(* IEC 61131-3 sources: STAR-PLC-Agent/results/raw/four_group_20261114/star_deepseek_v4/SELF011/generation/sim_00, 1 file *)

(* ---- test_program.st ---- *)
PROGRAM PLC_PRG
VAR
 BenchStep : UDINT := 0;
 BenchCalls : UDINT := 0;
 BenchDone : BOOL := FALSE;
 BenchUut0 : FB_Task;
 BenchUut1 : FB_Task;
 TraceIn_Start : ARRAY[0..12] OF BOOL;
 TraceIn_Stop : ARRAY[0..12] OF BOOL;
 TraceIn_Reset : ARRAY[0..12] OF BOOL;
 TraceIn_ExtendDone : ARRAY[0..12] OF BOOL;
 TraceIn_ClampDone : ARRAY[0..12] OF BOOL;
 TraceIn_ReleaseDone : ARRAY[0..12] OF BOOL;
 TraceIn_RetractDone : ARRAY[0..12] OF BOOL;
 TraceOut_Extend : ARRAY[0..12] OF BOOL;
 TraceOut_Clamp : ARRAY[0..12] OF BOOL;
 TraceOut_Release : ARRAY[0..12] OF BOOL;
 TraceOut_Retract : ARRAY[0..12] OF BOOL;
 TraceOut_Busy : ARRAY[0..12] OF BOOL;
 TraceOut_Done : ARRAY[0..12] OF BOOL;
END_VAR

IF NOT BenchDone THEN
 CASE BenchStep OF
 0:
   BenchUut0.Start := TRUE;
   BenchUut0.Stop := FALSE;
   BenchUut0.Reset := FALSE;
   BenchUut0.ExtendDone := FALSE;
   BenchUut0.ClampDone := FALSE;
   BenchUut0.ReleaseDone := FALSE;
   BenchUut0.RetractDone := TRUE;
   TraceIn_Start[0] := BenchUut0.Start;
   TraceIn_Stop[0] := BenchUut0.Stop;
   TraceIn_Reset[0] := BenchUut0.Reset;
   TraceIn_ExtendDone[0] := BenchUut0.ExtendDone;
   TraceIn_ClampDone[0] := BenchUut0.ClampDone;
   TraceIn_ReleaseDone[0] := BenchUut0.ReleaseDone;
   TraceIn_RetractDone[0] := BenchUut0.RetractDone;
   BenchUut0();
   TraceOut_Extend[0] := BenchUut0.Extend;
   TraceOut_Clamp[0] := BenchUut0.Clamp;
   TraceOut_Release[0] := BenchUut0.Release;
   TraceOut_Retract[0] := BenchUut0.Retract;
   TraceOut_Busy[0] := BenchUut0.Busy;
   TraceOut_Done[0] := BenchUut0.Done;
   BenchCalls := BenchCalls + 1;
 1:
   BenchUut0.Start := FALSE;
   BenchUut0.Stop := FALSE;
   BenchUut0.Reset := FALSE;
   BenchUut0.ExtendDone := TRUE;
   BenchUut0.ClampDone := FALSE;
   BenchUut0.ReleaseDone := FALSE;
   BenchUut0.RetractDone := FALSE;
   TraceIn_Start[1] := BenchUut0.Start;
   TraceIn_Stop[1] := BenchUut0.Stop;
   TraceIn_Reset[1] := BenchUut0.Reset;
   TraceIn_ExtendDone[1] := BenchUut0.ExtendDone;
   TraceIn_ClampDone[1] := BenchUut0.ClampDone;
   TraceIn_ReleaseDone[1] := BenchUut0.ReleaseDone;
   TraceIn_RetractDone[1] := BenchUut0.RetractDone;
   BenchUut0();
   TraceOut_Extend[1] := BenchUut0.Extend;
   TraceOut_Clamp[1] := BenchUut0.Clamp;
   TraceOut_Release[1] := BenchUut0.Release;
   TraceOut_Retract[1] := BenchUut0.Retract;
   TraceOut_Busy[1] := BenchUut0.Busy;
   TraceOut_Done[1] := BenchUut0.Done;
   BenchCalls := BenchCalls + 1;
 2:
   BenchUut0.Start := FALSE;
   BenchUut0.Stop := FALSE;
   BenchUut0.Reset := FALSE;
   BenchUut0.ExtendDone := FALSE;
   BenchUut0.ClampDone := TRUE;
   BenchUut0.ReleaseDone := FALSE;
   BenchUut0.RetractDone := FALSE;
   TraceIn_Start[2] := BenchUut0.Start;
   TraceIn_Stop[2] := BenchUut0.Stop;
   TraceIn_Reset[2] := BenchUut0.Reset;
   TraceIn_ExtendDone[2] := BenchUut0.ExtendDone;
   TraceIn_ClampDone[2] := BenchUut0.ClampDone;
   TraceIn_ReleaseDone[2] := BenchUut0.ReleaseDone;
   TraceIn_RetractDone[2] := BenchUut0.RetractDone;
   BenchUut0();
   TraceOut_Extend[2] := BenchUut0.Extend;
   TraceOut_Clamp[2] := BenchUut0.Clamp;
   TraceOut_Release[2] := BenchUut0.Release;
   TraceOut_Retract[2] := BenchUut0.Retract;
   TraceOut_Busy[2] := BenchUut0.Busy;
   TraceOut_Done[2] := BenchUut0.Done;
   BenchCalls := BenchCalls + 1;
 3:
   BenchUut0.Start := FALSE;
   BenchUut0.Stop := FALSE;
   BenchUut0.Reset := FALSE;
   BenchUut0.ExtendDone := FALSE;
   BenchUut0.ClampDone := FALSE;
   BenchUut0.ReleaseDone := TRUE;
   BenchUut0.RetractDone := FALSE;
   TraceIn_Start[3] := BenchUut0.Start;
   TraceIn_Stop[3] := BenchUut0.Stop;
   TraceIn_Reset[3] := BenchUut0.Reset;
   TraceIn_ExtendDone[3] := BenchUut0.ExtendDone;
   TraceIn_ClampDone[3] := BenchUut0.ClampDone;
   TraceIn_ReleaseDone[3] := BenchUut0.ReleaseDone;
   TraceIn_RetractDone[3] := BenchUut0.RetractDone;
   BenchUut0();
   TraceOut_Extend[3] := BenchUut0.Extend;
   TraceOut_Clamp[3] := BenchUut0.Clamp;
   TraceOut_Release[3] := BenchUut0.Release;
   TraceOut_Retract[3] := BenchUut0.Retract;
   TraceOut_Busy[3] := BenchUut0.Busy;
   TraceOut_Done[3] := BenchUut0.Done;
   BenchCalls := BenchCalls + 1;
 4:
   BenchUut0.Start := FALSE;
   BenchUut0.Stop := FALSE;
   BenchUut0.Reset := FALSE;
   BenchUut0.ExtendDone := FALSE;
   BenchUut0.ClampDone := FALSE;
   BenchUut0.ReleaseDone := FALSE;
   BenchUut0.RetractDone := TRUE;
   TraceIn_Start[4] := BenchUut0.Start;
   TraceIn_Stop[4] := BenchUut0.Stop;
   TraceIn_Reset[4] := BenchUut0.Reset;
   TraceIn_ExtendDone[4] := BenchUut0.ExtendDone;
   TraceIn_ClampDone[4] := BenchUut0.ClampDone;
   TraceIn_ReleaseDone[4] := BenchUut0.ReleaseDone;
   TraceIn_RetractDone[4] := BenchUut0.RetractDone;
   BenchUut0();
   TraceOut_Extend[4] := BenchUut0.Extend;
   TraceOut_Clamp[4] := BenchUut0.Clamp;
   TraceOut_Release[4] := BenchUut0.Release;
   TraceOut_Retract[4] := BenchUut0.Retract;
   TraceOut_Busy[4] := BenchUut0.Busy;
   TraceOut_Done[4] := BenchUut0.Done;
   BenchCalls := BenchCalls + 1;
 5:
   BenchUut0.Start := TRUE;
   BenchUut0.Stop := FALSE;
   BenchUut0.Reset := FALSE;
   BenchUut0.ExtendDone := FALSE;
   BenchUut0.ClampDone := FALSE;
   BenchUut0.ReleaseDone := FALSE;
   BenchUut0.RetractDone := TRUE;
   TraceIn_Start[5] := BenchUut0.Start;
   TraceIn_Stop[5] := BenchUut0.Stop;
   TraceIn_Reset[5] := BenchUut0.Reset;
   TraceIn_ExtendDone[5] := BenchUut0.ExtendDone;
   TraceIn_ClampDone[5] := BenchUut0.ClampDone;
   TraceIn_ReleaseDone[5] := BenchUut0.ReleaseDone;
   TraceIn_RetractDone[5] := BenchUut0.RetractDone;
   BenchUut0();
   TraceOut_Extend[5] := BenchUut0.Extend;
   TraceOut_Clamp[5] := BenchUut0.Clamp;
   TraceOut_Release[5] := BenchUut0.Release;
   TraceOut_Retract[5] := BenchUut0.Retract;
   TraceOut_Busy[5] := BenchUut0.Busy;
   TraceOut_Done[5] := BenchUut0.Done;
   BenchCalls := BenchCalls + 1;
 6:
   BenchUut1.Start := TRUE;
   BenchUut1.Stop := FALSE;
   BenchUut1.Reset := FALSE;
   BenchUut1.ExtendDone := FALSE;
   BenchUut1.ClampDone := FALSE;
   BenchUut1.ReleaseDone := FALSE;
   BenchUut1.RetractDone := FALSE;
   TraceIn_Start[6] := BenchUut1.Start;
   TraceIn_Stop[6] := BenchUut1.Stop;
   TraceIn_Reset[6] := BenchUut1.Reset;
   TraceIn_ExtendDone[6] := BenchUut1.ExtendDone;
   TraceIn_ClampDone[6] := BenchUut1.ClampDone;
   TraceIn_ReleaseDone[6] := BenchUut1.ReleaseDone;
   TraceIn_RetractDone[6] := BenchUut1.RetractDone;
   BenchUut1();
   TraceOut_Extend[6] := BenchUut1.Extend;
   TraceOut_Clamp[6] := BenchUut1.Clamp;
   TraceOut_Release[6] := BenchUut1.Release;
   TraceOut_Retract[6] := BenchUut1.Retract;
   TraceOut_Busy[6] := BenchUut1.Busy;
   TraceOut_Done[6] := BenchUut1.Done;
   BenchCalls := BenchCalls + 1;
 7:
   BenchUut1.Start := TRUE;
   BenchUut1.Stop := FALSE;
   BenchUut1.Reset := FALSE;
   BenchUut1.ExtendDone := FALSE;
   BenchUut1.ClampDone := FALSE;
   BenchUut1.ReleaseDone := FALSE;
   BenchUut1.RetractDone := TRUE;
   TraceIn_Start[7] := BenchUut1.Start;
   TraceIn_Stop[7] := BenchUut1.Stop;
   TraceIn_Reset[7] := BenchUut1.Reset;
   TraceIn_ExtendDone[7] := BenchUut1.ExtendDone;
   TraceIn_ClampDone[7] := BenchUut1.ClampDone;
   TraceIn_ReleaseDone[7] := BenchUut1.ReleaseDone;
   TraceIn_RetractDone[7] := BenchUut1.RetractDone;
   BenchUut1();
   TraceOut_Extend[7] := BenchUut1.Extend;
   TraceOut_Clamp[7] := BenchUut1.Clamp;
   TraceOut_Release[7] := BenchUut1.Release;
   TraceOut_Retract[7] := BenchUut1.Retract;
   TraceOut_Busy[7] := BenchUut1.Busy;
   TraceOut_Done[7] := BenchUut1.Done;
   BenchCalls := BenchCalls + 1;
 8:
   BenchUut1.Start := FALSE;
   BenchUut1.Stop := FALSE;
   BenchUut1.Reset := FALSE;
   BenchUut1.ExtendDone := TRUE;
   BenchUut1.ClampDone := FALSE;
   BenchUut1.ReleaseDone := FALSE;
   BenchUut1.RetractDone := FALSE;
   TraceIn_Start[8] := BenchUut1.Start;
   TraceIn_Stop[8] := BenchUut1.Stop;
   TraceIn_Reset[8] := BenchUut1.Reset;
   TraceIn_ExtendDone[8] := BenchUut1.ExtendDone;
   TraceIn_ClampDone[8] := BenchUut1.ClampDone;
   TraceIn_ReleaseDone[8] := BenchUut1.ReleaseDone;
   TraceIn_RetractDone[8] := BenchUut1.RetractDone;
   BenchUut1();
   TraceOut_Extend[8] := BenchUut1.Extend;
   TraceOut_Clamp[8] := BenchUut1.Clamp;
   TraceOut_Release[8] := BenchUut1.Release;
   TraceOut_Retract[8] := BenchUut1.Retract;
   TraceOut_Busy[8] := BenchUut1.Busy;
   TraceOut_Done[8] := BenchUut1.Done;
   BenchCalls := BenchCalls + 1;
 9:
   BenchUut1.Start := TRUE;
   BenchUut1.Stop := FALSE;
   BenchUut1.Reset := TRUE;
   BenchUut1.ExtendDone := FALSE;
   BenchUut1.ClampDone := TRUE;
   BenchUut1.ReleaseDone := FALSE;
   BenchUut1.RetractDone := FALSE;
   TraceIn_Start[9] := BenchUut1.Start;
   TraceIn_Stop[9] := BenchUut1.Stop;
   TraceIn_Reset[9] := BenchUut1.Reset;
   TraceIn_ExtendDone[9] := BenchUut1.ExtendDone;
   TraceIn_ClampDone[9] := BenchUut1.ClampDone;
   TraceIn_ReleaseDone[9] := BenchUut1.ReleaseDone;
   TraceIn_RetractDone[9] := BenchUut1.RetractDone;
   BenchUut1();
   TraceOut_Extend[9] := BenchUut1.Extend;
   TraceOut_Clamp[9] := BenchUut1.Clamp;
   TraceOut_Release[9] := BenchUut1.Release;
   TraceOut_Retract[9] := BenchUut1.Retract;
   TraceOut_Busy[9] := BenchUut1.Busy;
   TraceOut_Done[9] := BenchUut1.Done;
   BenchCalls := BenchCalls + 1;
 10:
   BenchUut1.Start := TRUE;
   BenchUut1.Stop := FALSE;
   BenchUut1.Reset := FALSE;
   BenchUut1.ExtendDone := FALSE;
   BenchUut1.ClampDone := FALSE;
   BenchUut1.ReleaseDone := FALSE;
   BenchUut1.RetractDone := TRUE;
   TraceIn_Start[10] := BenchUut1.Start;
   TraceIn_Stop[10] := BenchUut1.Stop;
   TraceIn_Reset[10] := BenchUut1.Reset;
   TraceIn_ExtendDone[10] := BenchUut1.ExtendDone;
   TraceIn_ClampDone[10] := BenchUut1.ClampDone;
   TraceIn_ReleaseDone[10] := BenchUut1.ReleaseDone;
   TraceIn_RetractDone[10] := BenchUut1.RetractDone;
   BenchUut1();
   TraceOut_Extend[10] := BenchUut1.Extend;
   TraceOut_Clamp[10] := BenchUut1.Clamp;
   TraceOut_Release[10] := BenchUut1.Release;
   TraceOut_Retract[10] := BenchUut1.Retract;
   TraceOut_Busy[10] := BenchUut1.Busy;
   TraceOut_Done[10] := BenchUut1.Done;
   BenchCalls := BenchCalls + 1;
 11:
   BenchUut1.Start := FALSE;
   BenchUut1.Stop := TRUE;
   BenchUut1.Reset := FALSE;
   BenchUut1.ExtendDone := TRUE;
   BenchUut1.ClampDone := FALSE;
   BenchUut1.ReleaseDone := FALSE;
   BenchUut1.RetractDone := FALSE;
   TraceIn_Start[11] := BenchUut1.Start;
   TraceIn_Stop[11] := BenchUut1.Stop;
   TraceIn_Reset[11] := BenchUut1.Reset;
   TraceIn_ExtendDone[11] := BenchUut1.ExtendDone;
   TraceIn_ClampDone[11] := BenchUut1.ClampDone;
   TraceIn_ReleaseDone[11] := BenchUut1.ReleaseDone;
   TraceIn_RetractDone[11] := BenchUut1.RetractDone;
   BenchUut1();
   TraceOut_Extend[11] := BenchUut1.Extend;
   TraceOut_Clamp[11] := BenchUut1.Clamp;
   TraceOut_Release[11] := BenchUut1.Release;
   TraceOut_Retract[11] := BenchUut1.Retract;
   TraceOut_Busy[11] := BenchUut1.Busy;
   TraceOut_Done[11] := BenchUut1.Done;
   BenchCalls := BenchCalls + 1;
 12:
   BenchUut1.Start := FALSE;
   BenchUut1.Stop := FALSE;
   BenchUut1.Reset := FALSE;
   BenchUut1.ExtendDone := FALSE;
   BenchUut1.ClampDone := FALSE;
   BenchUut1.ReleaseDone := FALSE;
   BenchUut1.RetractDone := FALSE;
   TraceIn_Start[12] := BenchUut1.Start;
   TraceIn_Stop[12] := BenchUut1.Stop;
   TraceIn_Reset[12] := BenchUut1.Reset;
   TraceIn_ExtendDone[12] := BenchUut1.ExtendDone;
   TraceIn_ClampDone[12] := BenchUut1.ClampDone;
   TraceIn_ReleaseDone[12] := BenchUut1.ReleaseDone;
   TraceIn_RetractDone[12] := BenchUut1.RetractDone;
   BenchUut1();
   TraceOut_Extend[12] := BenchUut1.Extend;
   TraceOut_Clamp[12] := BenchUut1.Clamp;
   TraceOut_Release[12] := BenchUut1.Release;
   TraceOut_Retract[12] := BenchUut1.Retract;
   TraceOut_Busy[12] := BenchUut1.Busy;
   TraceOut_Done[12] := BenchUut1.Done;
   BenchCalls := BenchCalls + 1;
 END_CASE;
 BenchStep := BenchStep + 1;
 IF BenchStep >= 13 THEN BenchDone := TRUE; END_IF;
END_IF;
END_PROGRAM
